(* IEC 61131-3 sources: plc-vscode/tests/st/test-ready/trust-platform/examples/OSCAT/shift_order_queue/non-oop/src, 3 files *)

(* ---- Configuration.st ---- *)
CONFIGURATION ShiftOrderQueueClassicConfiguration
RESOURCE Cpu0 ON PLC
    TASK MainTask (INTERVAL := T#100ms, PRIORITY := 1);
    PROGRAM Main WITH MainTask : Main;
END_RESOURCE
END_CONFIGURATION

(* ---- Main.st ---- *)
PROGRAM Main
VAR
    ShiftQueue : FIFO_16;
    NextShiftOrder : DWORD;
END_VAR

ShiftQueue(DIN := DWORD#16#3001, E := TRUE, RD := FALSE, WD := TRUE, RST := FALSE);
ShiftQueue(DIN := DWORD#16#3002, E := TRUE, RD := FALSE, WD := TRUE, RST := FALSE);
ShiftQueue(DIN := DWORD#0, E := TRUE, RD := TRUE, WD := FALSE, RST := FALSE);
NextShiftOrder := ShiftQueue.DOUT;
END_PROGRAM

(* ---- Tests.st ---- *)
TEST_PROGRAM ShiftOrderQueueClassicReturnsFirstOrderFirst
VAR
    ShiftQueue : FIFO_16;
END_VAR

ShiftQueue(DIN := DWORD#0, E := TRUE, RD := FALSE, WD := FALSE, RST := TRUE);
ShiftQueue(DIN := DWORD#16#3001, E := TRUE, RD := FALSE, WD := TRUE, RST := FALSE);
ShiftQueue(DIN := DWORD#16#3002, E := TRUE, RD := FALSE, WD := TRUE, RST := FALSE);
ShiftQueue(DIN := DWORD#0, E := TRUE, RD := TRUE, WD := FALSE, RST := FALSE);

ASSERT_EQUAL(EXPECTED := DWORD#16#3001, ACTUAL := ShiftQueue.DOUT);
END_TEST_PROGRAM
